Fanuc KAREL source: KT00311.KL

PROGRAM KT00311
%NOLOCKGROUP
VAR
  P1: POSITION
  P2: POSITION
  OUT: BOOLEAN
BEGIN
  OUT = P1 <> P2
END KT00311
